Fanuc KAREL source: KT00733.KL

PROGRAM KT00733
%NOLOCKGROUP
VAR
  ARG: ARRAY[4] OF REAL
  OUT: INTEGER
BEGIN
  OUT = ARRAY_LEN(ARG)
END KT00733
